TYPE ST_LightDefinition :
STRUCT
    sLocationCode : STRING(16);
    sLocationSlug : STRING(32);
    sLocationName : STRING(64);
    sId : STRING(32);
    sName : STRING(64);
    nButtonIndex : UINT;
END_STRUCT
END_TYPE

(* stored: Version 1.1.0.1
   DUT ST_LightDefinition: Id {f33452ad-55fc-49e6-bef5-f53ee005d41b} *)
